FUNCTION_BLOCK FB_Banddepalletizer IMPLEMENTS ITF_Banddepalletizer
VAR_INPUT
END_VAR
VAR_OUTPUT
END_VAR
VAR
END_VAR

{warning 'Add method implementation '}
METHOD Aborted : BOOL
END_METHOD

{warning 'Add method implementation '}
METHOD Aborting : BOOL
END_METHOD

{warning 'Add method implementation '}
METHOD Clearing : BOOL
END_METHOD

{warning 'Add method implementation '}
METHOD Execute : BOOL
END_METHOD

{warning 'Add method implementation '}
METHOD Held : BOOL
END_METHOD

{warning 'Add method implementation '}
METHOD Holding : BOOL
END_METHOD

{warning 'Add method implementation '}
METHOD Idle : BOOL
END_METHOD

{warning 'Add method implementation '}
METHOD Resetting : BOOL
END_METHOD

{warning 'Add method implementation '}
METHOD Starting : BOOL
END_METHOD

{warning 'Add method implementation '}
METHOD Stopped : BOOL
END_METHOD

{warning 'Add method implementation '}
METHOD Stopping : BOOL
END_METHOD

{warning 'Add method implementation '}
METHOD Suspended : BOOL
END_METHOD

{warning 'Add method implementation '}
METHOD Suspending : BOOL
END_METHOD

{warning 'Add method implementation '}
METHOD Unholding : BOOL
END_METHOD

{warning 'Add method implementation '}
METHOD Unsuspending : BOOL
END_METHOD

END_FUNCTION_BLOCK

(* stored: Version 1.1.0.1
   POU FB_Banddepalletizer: Id {dea9c50e-bcc0-4706-9e86-81f95655b873}, SpecialFunc None
   Folder Methods: Id {a781c065-e8ac-4b01-95ad-beaa1989158b}
   Method Aborted: Id {8a27e1f5-2cea-4c96-8327-4ebefd182309}
   Method Aborting: Id {500f5c57-804e-4edb-889d-3e65305c9d68}
   Method Clearing: Id {d947cecd-d02d-4310-9801-838a77815d3e}
   Method Execute: Id {b7667c93-f739-4270-8688-6ac20ba36ace}
   Method Held: Id {4a1acebb-e357-4258-b0d2-b79d3b5d6a54}
   Method Holding: Id {43996c19-55c1-4bfa-8f26-c5bbdb203676}
   Method Idle: Id {c8ec7455-f584-47b2-b053-5860a228cd72}
   Method Resetting: Id {d51a70a2-64f8-4fb1-bc27-1ff5c1562f4c}
   Method Starting: Id {356313a8-92a6-40b4-9b26-53e81edbd97a}
   Method Stopped: Id {a09bba40-f71e-4c0c-8a46-f2f883b49da7}
   Method Stopping: Id {c1f10999-dd62-4a90-beb9-88292f3ddd9e}
   Method Suspended: Id {039d7cfd-de79-4d03-aacd-36d334058b1c}
   Method Suspending: Id {9c691999-a116-487e-af04-a6b1e9db5be6}
   Method Unholding: Id {55845740-ad29-4a16-8d84-a5f3bb9cacbc}
   Method Unsuspending: Id {cf271d89-279e-4500-b8b2-cfde6201af80} *)
